(* IEC 61131-3 sources: pypi-mirror-400/packages/tc3tools/tc3tools-0.1.0.tar.gz/tc3tools-0.1.0/tests/fixtures/st, 19 files *)

(* ---- E_NodeStatus.st ---- *)
{attribute 'qualified_only'}
{attribute 'strict'}
TYPE E_NodeStatus :
(
    IDLE := 0,
    RUNNING,
    SUCCESS,
    FAILURE
) := IDLE;
END_TYPE

(* ---- E_Status.st ---- *)
{attribute 'qualified_only'}
{attribute 'strict'}
TYPE E_Status :
(
    Idle := 0,
    Initializing,
    Running,
    Paused,
    Stopping,
    Error := 99
) := Idle;
END_TYPE

(* ---- ST_Data.st ---- *)
TYPE ST_NestedData :
STRUCT
    bFlag : BOOL;
    nCount : INT;
END_STRUCT
END_TYPE

TYPE ST_Data :
STRUCT
    nId : UDINT;
    sName : STRING(80);
    fValue : REAL;
    dtTimestamp : DT;
    aBuffer : ARRAY[0..255] OF BYTE;
    stNested : ST_NestedData;
END_STRUCT
END_TYPE

(* ---- GVL_Constants.st ---- *)
{attribute 'qualified_only'}
VAR_GLOBAL CONSTANT
    GC_VERSION : STRING := '1.0.0';
    GC_MAX_DEVICES : UINT := 64;
    GC_TIMEOUT_MS : TIME := T#5000MS;
    GC_PI : LREAL := 3.14159265358979;
END_VAR

VAR_GLOBAL
    g_bSystemReady : BOOL;
    g_nActiveDevices : UINT;
END_VAR

VAR_GLOBAL RETAIN
    g_nTotalCycles : ULINT;
    g_dtLastRun : DT;
END_VAR

(* ---- I_Device.st ---- *)
INTERFACE I_Device

PROPERTY DeviceId : UDINT
END_PROPERTY

PROPERTY IsOnline : BOOL
END_PROPERTY

METHOD Initialize : BOOL
VAR_INPUT
    nId : UDINT;
END_VAR
END_METHOD

METHOD Execute : BOOL
END_METHOD

METHOD GetStatus : INT
END_METHOD

END_INTERFACE

(* ---- I_Errorable.st ---- *)
INTERFACE I_Errorable

    METHOD HasError : BOOL
    END_METHOD

    METHOD GetError : ST_Error
    END_METHOD

    METHOD ClearError
    END_METHOD

END_INTERFACE

(* ---- I_TreeNode.st ---- *)
INTERFACE I_TreeNode

    // Method: Tick - Main execution method
    METHOD Tick : E_NodeStatus
    END_METHOD

    // Method: Halt - Stop execution
    METHOD Halt
    END_METHOD

    // Method: Reset - Reset state
    METHOD Reset : BOOL
    END_METHOD

    // Method: GetPath - Get node path
    METHOD GetPath : STRING(255)
    END_METHOD

    // Method: GetNodeName - Get node name
    METHOD GetNodeName : STRING(50)
    END_METHOD

    // Method: SetParent - Set parent node
    METHOD SetParent
        VAR_INPUT
            ipParent : I_TreeNode;
        END_VAR
    END_METHOD

    // Method: GetProgress - Get progress value
    METHOD GetProgress : REAL
    END_METHOD

    // Error handling methods
    METHOD HasError : BOOL
    END_METHOD

    METHOD GetError : ST_Error
    END_METHOD

    METHOD ClearError
    END_METHOD

END_INTERFACE

(* ---- FC_Calculate.st ---- *)
FUNCTION FC_Calculate : REAL
VAR_INPUT
    fA : REAL;
    fB : REAL;
    eOperation : INT;
END_VAR
VAR
    fResult : REAL;
END_VAR

CASE eOperation OF
    0:
        fResult := fA + fB;
    1:
        fResult := fA - fB;
    2:
        fResult := fA * fB;
    3:
        IF fB <> 0.0 THEN
            fResult := fA / fB;
        ELSE
            fResult := 0.0;
        END_IF
ELSE
    fResult := 0.0;
END_CASE

FC_Calculate := fResult;

END_FUNCTION

(* ---- FB_ActionNode.st ---- *)
(* Action node that extends base node *)
FUNCTION_BLOCK FB_ActionNode EXTENDS FB_BaseNode
VAR
    _nExecutionCount : INT;
    _bFirstExecution : BOOL := TRUE;
END_VAR

METHOD Tick : E_NodeStatus
    IF _bFirstExecution THEN
        _bFirstExecution := FALSE;
        _nExecutionCount := 0;
    END_IF

    _nExecutionCount := _nExecutionCount + 1;

    IF HasError() THEN
        Tick := E_NodeStatus.FAILURE;
    ELSE
        Tick := E_NodeStatus.SUCCESS;
    END_IF

    eLastStatus := Tick;
END_METHOD

METHOD Reset : BOOL
    SUPER^.Reset();
    _nExecutionCount := 0;
    _bFirstExecution := TRUE;
    Reset := TRUE;
END_METHOD

METHOD PUBLIC GetExecutionCount : INT
    GetExecutionCount := _nExecutionCount;
END_METHOD

END_FUNCTION_BLOCK

(* ---- FB_AlwaysFailure.st ---- *)
(* Simple derived node - always returns FAILURE *)
FUNCTION_BLOCK FB_AlwaysFailure EXTENDS FB_BaseNode

METHOD Tick : E_NodeStatus
    Tick := E_NodeStatus.FAILURE;
    eLastStatus := E_NodeStatus.FAILURE;
END_METHOD

END_FUNCTION_BLOCK

(* ---- FB_AlwaysSuccess.st ---- *)
(* Simple derived node - always returns SUCCESS *)
FUNCTION_BLOCK FB_AlwaysSuccess EXTENDS FB_BaseNode

METHOD Tick : E_NodeStatus
    Tick := E_NodeStatus.SUCCESS;
    eLastStatus := E_NodeStatus.SUCCESS;
    SetProgressComplete();
END_METHOD

END_FUNCTION_BLOCK

(* ---- FB_BaseNode.st ---- *)
{attribute 'qualified_only'}
FUNCTION_BLOCK FB_BaseNode IMPLEMENTS I_TreeNode, I_Errorable
VAR
    eLastStatus : E_NodeStatus := E_NodeStatus.IDLE;
    _sNodeName : STRING(50);
    rProgress : REAL := 0.0;
    _fbErrorHandler : FB_ErrorHandler;
    _sFailedChildName : STRING(50);
    _ipParent : I_TreeNode;
    _bHalted : BOOL := FALSE;
END_VAR

PROPERTY NodeName : STRING(50)
    GET
    NodeName := _sNodeName;
    END_GET
    SET
    _sNodeName := NodeName;
    _fbErrorHandler.Initialize(_sNodeName);
    END_SET
END_PROPERTY

METHOD Tick : E_NodeStatus
    Tick := E_NodeStatus.IDLE;
END_METHOD

METHOD Halt
    _bHalted := TRUE;
    eLastStatus := E_NodeStatus.IDLE;
    rProgress := 0.0;
END_METHOD

METHOD Reset : BOOL
    _bHalted := FALSE;
    eLastStatus := E_NodeStatus.IDLE;
    rProgress := 0.0;
    ClearError();
    Reset := TRUE;
END_METHOD

METHOD PUBLIC SetParent
    VAR_INPUT
        ipParent : I_TreeNode;
    END_VAR
    _ipParent := ipParent;
END_METHOD

METHOD PUBLIC GetPath : STRING(255)
    VAR
        sPath : STRING(255);
    END_VAR
    IF _ipParent <> 0 THEN
        sPath := _ipParent.GetPath();
        IF LEN(sPath) > 0 THEN
            sPath := CONCAT(sPath, '/');
        END_IF
        sPath := CONCAT(sPath, _sNodeName);
    ELSE
        sPath := _sNodeName;
    END_IF
    GetPath := sPath;
END_METHOD

METHOD PUBLIC GetNodeName : STRING(50)
    GetNodeName := _sNodeName;
END_METHOD

METHOD PUBLIC SetError
    VAR_INPUT
        eErrorId : E_ErrorId;
        sMessage : STRING(255);
    END_VAR
    _fbErrorHandler.Raise(eErrorId, sMessage);
END_METHOD

METHOD PUBLIC HasError : BOOL
    HasError := _fbErrorHandler.IsActive();
END_METHOD

METHOD PUBLIC GetError : ST_Error
    GetError := _fbErrorHandler.GetError();
END_METHOD

METHOD PUBLIC ClearError
    _fbErrorHandler.Clear();
    _sFailedChildName := '';
END_METHOD

METHOD PUBLIC GetProgress : REAL
    GetProgress := rProgress;
END_METHOD

METHOD PROTECTED UpdateProgress
    VAR_INPUT
        nCurrent : INT;
        nTotal : INT;
    END_VAR
    IF nTotal > 0 THEN
        rProgress := (INT_TO_REAL(nCurrent) / INT_TO_REAL(nTotal)) * 100.0;
    ELSE
        rProgress := 0.0;
    END_IF
END_METHOD

METHOD PROTECTED SetProgressComplete
    rProgress := 100.0;
END_METHOD

END_FUNCTION_BLOCK

(* ---- FB_ConditionNode.st ---- *)
{attribute 'qualified_only'}
{attribute 'strict'}
(* Condition node with EXTENDS and multiple interface check *)
FUNCTION_BLOCK FB_ConditionNode EXTENDS FB_BaseNode
VAR_INPUT
    bCondition : BOOL;
END_VAR
VAR
    _bLastCondition : BOOL;
    _nEvaluationCount : UDINT;
END_VAR

METHOD Tick : E_NodeStatus
    _nEvaluationCount := _nEvaluationCount + 1;
    _bLastCondition := bCondition;

    IF bCondition THEN
        Tick := E_NodeStatus.SUCCESS;
        SetProgressComplete();
    ELSE
        Tick := E_NodeStatus.FAILURE;
    END_IF

    eLastStatus := Tick;
END_METHOD

METHOD Reset : BOOL
    SUPER^.Reset();
    _bLastCondition := FALSE;
    _nEvaluationCount := 0;
    Reset := TRUE;
END_METHOD

PROPERTY EvaluationCount : UDINT
    GET
    EvaluationCount := _nEvaluationCount;
    END_GET
END_PROPERTY

PROPERTY LastCondition : BOOL
    GET
    LastCondition := _bLastCondition;
    END_GET
END_PROPERTY

END_FUNCTION_BLOCK

(* ---- FB_EdgeCases.st ---- *)
{attribute 'reflection'}
{attribute 'hide_all_locals'}
FUNCTION_BLOCK FB_EdgeCases EXTENDS FB_Base IMPLEMENTS I_Device
VAR_INPUT
    {attribute 'OPC.UA.DA' := '1'}
    fSetpoint : REAL := 0.0;
    sDescription : STRING(255) := 'Default description';
END_VAR
VAR_OUTPUT
    {attribute 'OPC.UA.DA.Access' := '1'}
    fActualValue : REAL;
END_VAR
VAR CONSTANT
    C_MAX_VALUE : REAL := 100.0;
    C_MIN_VALUE : REAL := -100.0;
END_VAR
VAR
    // Single line comment
    _state : INT;
    (* Block comment *)
    _timer : TON;
    (*
        Multi-line
        block comment
    *)
    _lastValue : REAL;
END_VAR

// Edge case: IF-ELSIF-ELSE chain
IF fSetpoint > C_MAX_VALUE THEN
    fActualValue := C_MAX_VALUE;
ELSIF fSetpoint < C_MIN_VALUE THEN
    fActualValue := C_MIN_VALUE;
ELSIF fSetpoint = 0.0 THEN
    fActualValue := _lastValue;
ELSE
    fActualValue := fSetpoint;
END_IF

// Edge case: Nested IF
IF _state = 1 THEN
    IF fSetpoint > 0.0 THEN
        IF _timer.Q THEN
            fActualValue := fSetpoint;
        END_IF
    END_IF
END_IF

// Edge case: WHILE loop
WHILE _state = 0 DO
    _state := 1;
END_WHILE

// Edge case: REPEAT-UNTIL
REPEAT
    _lastValue := fActualValue;
UNTIL _state <> 1
END_REPEAT

_lastValue := fActualValue;

METHOD PUBLIC FB_init : BOOL
VAR_INPUT
    bInitRetains : BOOL;
    bInCopyCode : BOOL;
END_VAR
    _state := 0;
    FB_init := TRUE;
END_METHOD

{attribute 'TcRpcEnable'}
METHOD ProcessData : BOOL
VAR_INPUT
    nSize : UDINT;
END_VAR
VAR
    i : UDINT;
END_VAR
    FOR i := 0 TO nSize - 1 DO
        // Process each item
        _lastValue := _lastValue + 1.0;
    END_FOR
    ProcessData := TRUE;
END_METHOD

END_FUNCTION_BLOCK

(* ---- FB_Sample.st ---- *)
FUNCTION_BLOCK FB_Sample
VAR_INPUT
    bEnable : BOOL;
    nValue : INT;
END_VAR
VAR_OUTPUT
    bDone : BOOL;
    nResult : INT;
END_VAR
VAR
    _state : INT;
END_VAR

IF bEnable THEN
    _state := _state + 1;
    nResult := nValue * 2;
    bDone := TRUE;
ELSE
    bDone := FALSE;
END_IF
END_FUNCTION_BLOCK

(* ---- FB_SimpleBlock.st ---- *)
FUNCTION_BLOCK FB_SimpleBlock
VAR_INPUT
    bEnable : BOOL;
    nValue : INT;
END_VAR
VAR_OUTPUT
    bDone : BOOL;
    nResult : INT;
END_VAR
VAR
    _state : INT;
END_VAR

IF bEnable THEN
    nResult := nValue * 2;
    bDone := TRUE;
ELSE
    bDone := FALSE;
END_IF

END_FUNCTION_BLOCK

(* ---- FB_WithMethods.st ---- *)
{attribute 'qualified_only'}
{attribute 'strict'}
FUNCTION_BLOCK FB_WithMethods
VAR_INPUT
    bExecute : BOOL;
END_VAR
VAR_OUTPUT
    bBusy : BOOL;
    bError : BOOL;
    nErrorId : UDINT;
END_VAR
VAR
    _counter : INT;
    _initialized : BOOL;
END_VAR

(* Main implementation *)
IF bExecute AND NOT _initialized THEN
    Initialize();
END_IF

METHOD PUBLIC Initialize : BOOL
VAR_INPUT
    nStartValue : INT := 0;
END_VAR
VAR
    i : INT;
END_VAR
    FOR i := 0 TO 10 DO
        _counter := _counter + 1;
    END_FOR
    _initialized := TRUE;
    Initialize := TRUE;
END_METHOD

METHOD PRIVATE Reset
VAR
    temp : INT;
END_VAR
    _counter := 0;
    _initialized := FALSE;
END_METHOD

METHOD Calculate : REAL
VAR_INPUT
    fInput : REAL;
END_VAR
VAR_OUTPUT
    fOutput : REAL;
END_VAR
VAR
    fTemp : REAL;
END_VAR
    CASE _counter OF
        0:
            fTemp := 0.0;
        1..5:
            fTemp := fInput * 2.0;
        6, 7, 8:
            fTemp := fInput / 2.0;
    ELSE
        fTemp := fInput;
    END_CASE

    fOutput := fTemp;
    Calculate := fTemp;
END_METHOD

END_FUNCTION_BLOCK

(* ---- FB_WithProperties.st ---- *)
FUNCTION_BLOCK FB_WithProperties
VAR
    _value : INT;
    _name : STRING(80);
    _enabled : BOOL;
END_VAR

PROPERTY PUBLIC Value : INT
GET
VAR
    temp : INT;
END_VAR
    temp := _value;
    Value := temp;
END_GET
SET
    _value := Value;
END_SET
END_PROPERTY

PROPERTY Name : STRING(80)
GET
    Name := _name;
END_GET
SET
    _name := Name;
END_SET
END_PROPERTY

PROPERTY Enabled : BOOL
GET
    Enabled := _enabled;
END_GET
END_PROPERTY

METHOD DoWork : BOOL
    IF _enabled THEN
        _value := _value + 1;
        DoWork := TRUE;
    END_IF
END_METHOD

END_FUNCTION_BLOCK

(* ---- PRG_Main.st ---- *)
PROGRAM PRG_Main
VAR
    fbSimple : FB_SimpleBlock;
    fbMethods : FB_WithMethods;
    bStart : BOOL;
    nCycleCount : UDINT;
END_VAR

nCycleCount := nCycleCount + 1;

fbSimple(
    bEnable := bStart,
    nValue := 42
);

IF fbSimple.bDone THEN
    fbMethods(bExecute := TRUE);
END_IF

END_PROGRAM
